(* IEC 61131-3 sources: openplc-editor-canopen/src/backend/shared/transpilers/st-transpiler/__tests__/fixtures/ld-relayout-corpus/ld-corpus-imported/expected-st, 4 files *)

(* ---- _project.st ---- *)
CONFIGURATION Config0

  RESOURCE Res0 ON PLC
    TASK task0(INTERVAL := T#20ms,PRIORITY := 1);
    PROGRAM instance0 WITH task0 : main;
  END_RESOURCE
END_CONFIGURATION

(* ---- main_fbd.st ---- *)
PROGRAM main_fbd
  VAR
    TON5 : TON;
    TON6 : TON;
    TON7 : TON;
  END_VAR

  TON5();
  TON6();
  TON7();
  TON7();
END_PROGRAM

(* ---- main_ld.st ---- *)
PROGRAM main_ld
  VAR
    man_mode : BOOL;
    Moisture : BOOL;
    timeout : BOOL;
    run_valve : BOOL;
    new_ct : BOOL;
    T_Max : TIME;
    test_something : INT;
    TON0 : TON;
    TOF0 : TOF;
    CTU0 : CTU;
  END_VAR

  run_valve := NOT(TOF0.Q) AND Moisture AND NOT(man_mode);
  TON0(IN := run_valve, PT := T_Max);
  TOF0(IN := TON0.Q, PT := T_Max);
  timeout := TOF0.Q;
  CTU0(CU := new_ct, R := NOT(man_mode), PV := 10);
  test_something := CTU0.CV;
END_PROGRAM

(* ---- motor_ladder.st ---- *)
PROGRAM motor_ladder

  Lamp := Motor;
END_PROGRAM
